(* IEC 61131-3 sources: moqui-plc/iec61131/moqui/framework/src/test/robot-arm, 1 file *)

(* ---- TestRobotArmPlanning.st ---- *)
PROGRAM TestRobotArmPlanning

	;
	(* The planning task must have a cycle that is exactly N×T_bus with N integers.
	 * If the values ​​do not meet this constraint, CODESYS calculates an inconsistent CP configuration and each MC_MoveLinearAbsolute fails.
	 *)
	END_PROGRAM
